Fanuc KAREL source: KA00021.KL

PROGRAM KA00021
%NOLOCKGROUP
VAR
  SRC: REAL
  DST: VECTOR
BEGIN
  SRC = 2.0
  DST = SRC
END KA00021
